FUNCTION_BLOCK FB_Generic
VAR_GENERIC CONSTANT
	nMax : DINT := 10;
END_VAR IMPLEMENTS I_Collection, I_Enumerator;
VAR
	aItems : ARRAY[0..nMax] OF INT;
END_VAR

aItems[0] := 1;

END_FUNCTION_BLOCK

(* stored: Version 1.1.0.1, ProductVersion 3.1.4026.12
   POU FB_Generic: Id {11111111-2222-3333-4444-666666666666}, SpecialFunc None *)
